// TwinCAT 3 PLC project plc
// ProgramVersion: 3.1.4026.24
// libraries:
//   Tc2_Standard, * (Beckhoff Automation GmbH)
//   Tc2_System, * (Beckhoff Automation GmbH)
//   Tc3_Database, * (Beckhoff Automation GmbH)
// project tree:
//   DUTs/ ST_Signals.TcDUT
//   / PlcTask.TcTTO
//   POUs/ E_FunctionType.TcDUT, FB_FunctionGenerator.TcPOU, MAIN.TcPOU
// real-time tasks:
//   TASK PlcTask: cycle T#10ms, priority 20, ADS port 350

CONFIGURATION plc
    RESOURCE PLC ON TwinCAT3
        TASK PlcTask(INTERVAL := T#10ms, PRIORITY := 20);
        PROGRAM MAIN WITH PlcTask : MAIN;
    END_RESOURCE
END_CONFIGURATION

// ---- DUTs/ST_Signals.TcDUT
TYPE ST_Signals :
STRUCT
    {attribute 'TagName' := 'ID'}
    signal : STRING(255);
    
    {attribute 'FieldName' := 'Value'}
    value : LREAL := -1;
	
END_STRUCT
END_TYPE

// ---- POUs/E_FunctionType.TcDUT
TYPE E_FunctionType :
(
	eSine,
	eSquare,
	ePulse,
	eTriangular,
	eSawtooth,	
	eAM
);
END_TYPE

// ---- POUs/MAIN.TcPOU
PROGRAM MAIN
VAR
	fbSignalSaw				: FB_FunctionGenerator;
	rSignal1				: LREAL;		// Señal dientes de sierra generada por plc
	fbSignalSinus1			: FB_FunctionGenerator;
	rSignal2				: LREAL;		// Señal senoidal generada por plc
	fbDBAutoLog				: FB_PLCDBAutoLogEvt(sNetID:='', tTimeout:=T#5S);
	bAutoLogStart			: BOOL;
	bErrAutoLog				: BOOL;
	aAutoLogStatus			: ARRAY [1..1] OF ST_AutoLogGrpStatus;		// Estado de la conexion Autolog con la DB
	rTrig1					: R_TRIG;
	fTrig2					: F_TRIG;
	bRun					: BOOL;			// Arranca DB Autolog
	bStop					: BOOL;			// Detiene DB Autolog
	timerReset				: TON;
	bErrorInfluxdb			: BOOL;			// Error en la conexion con la DB
	iReconexiones			: INT;			// Contador de reintentos de conexion con la DB
END_VAR

fbSignalSaw(
	bEnable:= TRUE, 
	fFrequency:= 0.2, 
	fAmplitude:= 10, 
	fOffset:= 0, 
	nDutyCycle:= , 
	eFunction:= E_FunctionType.eSawtooth, 
	rSignal:= rSignal1, 
	bError=> );
	
fbSignalSinus1(
	bEnable:= TRUE, 
	fFrequency:= 0.1, 
	fAmplitude:= 5, 
	fOffset:= 0, 
	nDutyCycle:= , 
	eFunction:= E_FunctionType.eSine, 
	rSignal:= rSignal2, 
	bError=> );

rTrig1(CLK:=bAutoLogStart, Q=> );
fTrig2(CLK:=bAutoLogStart, Q=> );

IF _TaskInfo[1].FirstCycle THEN
	bAutoLogStart := TRUE;  // No se inicializa la variable en la declaracion ya que el bloque trigger no detectaría el cambio
END_IF

// Se usa la salida trigger para generar el mensaje en el log, que solo necesita 1 ciclo
// La activacion del autolog con el método Start() tarda unos ciclos
IF rTrig1.Q THEN
	ADSLOGSTR(msgCtrlMask:= ADSLOG_MSGTYPE_WARN OR ADSLOG_MSGTYPE_LOG, msgFmtStr:= 'Autolog Started %s', strArg:='' );
	bRun := TRUE;
END_IF

IF fTrig2.Q THEN
	ADSLOGSTR(msgCtrlMask:= ADSLOG_MSGTYPE_WARN OR ADSLOG_MSGTYPE_LOG, msgFmtStr:= 'Autolog Stopped %s', strArg:='' );
	bStop := TRUE;
END_IF

IF bRun THEN
	IF fbDBAutoLog.Start() THEN
		bRun := FALSE;
	END_IF
END_IF

// EL método Stop también necesita varios ciclos
IF bStop THEN
	IF fbDBAutoLog.Stop() THEN
		bStop := FALSE;
	END_IF
END_IF

// El método de diagnóstico se puede ejecutar cíclicamente
IF bAutoLogStart THEN
	aAutoLogStatus[1].hAutoLogGrpID := 3;
	fbDBAutoLog.Status(tCheckCycle:=T#3S , pError:=ADR(bErrAutoLog) , pAutoLogGrpStatus:=ADR(aAutoLogStatus) , cbAutoLogGrpStatus:=SIZEOF(aAutologStatus) );
	// Si devuelve aAutoLogStatus[1].hrErrorCode= 16#989103E8 la base de datos InfluxDB está detenida
	IF NOT fbDBAutoLog.bBusy_Status THEN
		bErrorInfluxdb := aAutoLogStatus[1].bError;
	END_IF
END_IF

// En caso de error en la conexion con InfluxDB, resetea la funcion autolog cada 3s y comprueba la conexion 
IF bErrorInfluxdb THEN
	bAutoLogStart := FALSE;
	timerReset(IN:=TRUE , PT:=T#3S);
	IF timerReset.Q THEN
		bAutoLogStart := TRUE;
		IF NOT fbDBAutoLog.bBusy_Status THEN
			iReconexiones := iReconexiones+1;
			timerReset(IN:=FALSE);
			bErrorInfluxdb := aAutoLogStatus[1].bError;
		END_IF
	END_IF
ELSE
	timerReset(IN:=FALSE);	
END_IF

END_PROGRAM

// ---- POUs/FB_FunctionGenerator.TcPOU
// Generates a signal build up by the specified function type. v1.2
FUNCTION_BLOCK FB_FunctionGenerator
VAR_INPUT
	bEnable		: BOOL := TRUE;
	fFrequency	: LREAL := 1000;	// in [Hz]
	fAmplitude	: LREAL := 1;
	fOffset		: LREAL;
	nDutyCycle	: UINT := 50;		// % (for pulse function)
	eFunction	: E_FunctionType := E_FunctionType.eSine;	//Default sine wave
END_VAR
VAR_IN_OUT
	rSignal		: LREAL;			//output signal
END_VAR
VAR_OUTPUT
	bError		: BOOL;
END_VAR

VAR
	bInit						: BOOL := TRUE;
	fbGetTaskIdx				: GETCURTASKINDEX;
	
	fLastFrequency				: LREAL;		// in [Hz]
	fLastAmplitude				: LREAL;
	fLastOffset					: LREAL;
	nLastDutyCycle				: UINT;
	eLastFunction				: E_FunctionType;
	
//	nSamples					: UDINT;
	fCycleTime					: LREAL;		// in [s]
	fDelta						: LREAL;		// amplitude delta per sample
	fPhase						: LREAL;		// in [°]
	nSign						: INT := 1;		// 1 or -1
	fLastSignalValue			: LREAL;		// amplitude
	fPeriod						: LREAL;		// in [s]
	fAngularIncrement			: LREAL;		// in [°]
	fAngularIncrementPerCycle	: LREAL;		// in [°]
	fAngularIncrementPerSample	: LREAL;		// in [°]
	(* for modulated signal *)
	fCarrierFrequency			: LREAL := 500;	// in [Hz] (sine)
	fCarrierAmplitude			: LREAL := 1;
	fCarrierPeriod				: LREAL;		// in [s]
	fCarrierAngularIncrement			: LREAL;		// in [°]
	fCarrierAngularIncrementPerCycle	: LREAL;		// in [°]
//	fCarrierAngularIncrementPerSample	: LREAL;		// in [°]
END_VAR

IF bEnable THEN
	IF fLastFrequency <> fFrequency THEN
		bInit := TRUE; // For automatic initializing
		fLastFrequency := fFrequency;
	END_IF
	IF fLastAmplitude <> fAmplitude THEN
		bInit := TRUE; // For automatic initializing
		fLastAmplitude := fAmplitude;
	END_IF
	IF fLastOffset <> fOffset THEN
		bInit := TRUE; // For automatic initializing
		fLastOffset := fOffset;
	END_IF
	IF nLastDutyCycle <> nDutyCycle THEN
		bInit := TRUE; // For automatic initializing
		nLastDutyCycle := nDutyCycle;
	END_IF
	IF eLastFunction <> eFunction THEN
		bInit := TRUE; // For automatic initializing
		eLastFunction := eFunction;
	END_IF
	IF bInit THEN
		// Get taks info	
		fbGetTaskIdx();
		fCycleTime := TwinCAT_SystemInfoVarList._TaskInfo[fbGetTaskIdx.index].CycleTime (*100ns*) / (10.0 * 1000.0 * 1000.0);	
		fLastSignalValue := 0;
		nSign := 1;
		fAngularIncrement := 0;
		// Flush out old data
		MEMSET(ADR(rSignal), 0, SIZEOF(rSignal));
		IF fFrequency <> 0 AND fCycleTime > 0 THEN		
			// Calculate period, increments per plc cycle, increment per oversample

			IF eFunction = E_FunctionType.eSine THEN
				fPeriod := 1/fFrequency;
				fAngularIncrementPerCycle := 360*(fCycleTime/fPeriod);
				// no phase adjustment
				bInit := FALSE;	
			ELSIF eFunction = E_FunctionType.eSquare	THEN
				fPeriod := 1/fFrequency;
				fAngularIncrementPerCycle  := 360*(fCycleTime/fPeriod);
				fPhase := 0.5*360;
				bInit := FALSE;
			ELSIF eFunction = E_FunctionType.ePulse THEN
				fPeriod := 1/fFrequency;
				fAngularIncrementPerCycle  := 360*(fCycleTime/fPeriod);
				IF nDutyCycle > 100 THEN
					nDutyCycle := 100;
				END_IF
				fPhase := (UDINT_TO_LREAL(nDutyCycle)/100)*360;
				bInit := FALSE;					
			ELSIF eFunction = E_FunctionType.eTriangular THEN
				fPeriod := 1/fFrequency;				
				fAngularIncrementPerCycle  := 360*(fCycleTime/fPeriod);
				fAngularIncrementPerSample := fAngularIncrementPerCycle;
				fPhase := 0.5*360; 
				fDelta := 4*(fAmplitude/(360/fAngularIncrementPerSample));				
				bInit := FALSE;
			ELSIF eFunction = E_FunctionType.eSawtooth THEN
				fPeriod := 1/fFrequency;			
				fAngularIncrementPerCycle  := 360*(fCycleTime/fPeriod);		
				fAngularIncrementPerSample := fAngularIncrementPerCycle;
				fDelta := fAmplitude/(360/fAngularIncrementPerSample);
				bInit := FALSE;
			ELSIF eFunction = E_FunctionType.eAM THEN
				fPeriod := 1/fFrequency;
				fAngularIncrementPerCycle := 360*(fCycleTime/fPeriod);
				// no phase adjustment
				fCarrierPeriod := 1/fCarrierFrequency;
				fCarrierAngularIncrementPerCycle := 360*(fCycleTime/fCarrierPeriod);
				// no phase adjustment	
				bInit := FALSE;			
			ELSE
				bError := TRUE;	
			END_IF
		ELSE
			bError := TRUE;
		END_IF
	END_IF
	
	// Enable function generator
	IF NOT bError THEN		
		CASE eFunction OF		
			// sine: typical for vibrations originating from rotating machine
			E_FunctionType.eSine: Sine();
			
			// square: mixed sine signals good for analyzing spectrum				
			E_FunctionType.eSquare: Square();
			
			// pulse: mixed sine signals good for analyzing spectrum				
			E_FunctionType.ePulse: Pulse();
	
			// sawtooth: ramp-type vibrations, continuously increasing			
			E_FunctionType.eSawtooth: Sawtooth();
		
			// triangular: mixed sine signals good for analyzing spectrum
			E_FunctionType.eTriangular: Triangular();
		
			// amplitude modulation: typical for vibrations originating from gear-tooth failure or bearing faults
			// Carrier signal with own frequency and amplitude		
			E_FunctionType.eAM: AM();			
		END_CASE
	END_IF
ELSE
	// Flush out old data
	MEMSET(ADR(rSignal), 0, SIZEOF(rSignal));
END_IF

METHOD PRIVATE AM
VAR_INPUT
END_VAR
// base signal * carrier signal
rSignal:= ( fAmplitude*SIN(2*PI*(fAngularIncrement)/360) + fOffset )
						* ( fCarrierAmplitude*SIN(2*PI*(fCarrierAngularIncrement)/360) );

// Increment angular positions
fAngularIncrement := fAngularIncrement + fAngularIncrementPerCycle;
fCarrierAngularIncrement := fCarrierAngularIncrement + fCarrierAngularIncrementPerCycle;
END_METHOD

METHOD PRIVATE Pulse
VAR_INPUT
END_VAR
// For pulse wave (unequal phases)
IF (fAngularIncrement >= 360) THEN
	fAngularIncrement := fAngularIncrement - DINT_TO_LREAL(LREAL_TO_DINT(fAngularIncrement/360))*360;
	// or with Tc2_Math library: fAngularIncrement := LMOD(fAngularIncrement,360);
END_IF
IF (fAngularIncrement < fPhase) THEN
	nSign := 1;		
ELSIF (fAngularIncrement >= fPhase) THEN
	nSign := 0;
END_IF

rSignal:= nSign*fAmplitude;

rSignal:= rSignal+ fOffset;
END_METHOD

METHOD PRIVATE Sawtooth
VAR_INPUT
END_VAR

// For sawtooth wave (equal phase = period/2)
IF (fAngularIncrement >= 360) THEN
	fAngularIncrement := fAngularIncrement - DINT_TO_LREAL(LREAL_TO_DINT(fAngularIncrement/360))*360;
	// or with Tc2_Math library: fAngularIncrement := LMOD(fAngularIncrement,360);
	fLastSignalValue := fLastSignalValue -fAmplitude;
END_IF
fAngularIncrement := fAngularIncrement + fAngularIncrementPerSample;

rSignal:= fLastSignalValue + fDelta;

// Store last sample
fLastSignalValue := rSignal;

rSignal:= rSignal+ fOffset;
END_METHOD

METHOD PRIVATE Sine
VAR_INPUT
END_VAR

rSignal := fAmplitude*SIN(2*PI*(fAngularIncrement/360));

rSignal := rSignal + fOffset;


// Increment angular position
fAngularIncrement := fAngularIncrement + fAngularIncrementPerCycle;
END_METHOD

METHOD PRIVATE Square
VAR_INPUT
END_VAR

// For square wave (equal phase = period/2)
IF (fAngularIncrement >= 360) THEN
	fAngularIncrement := fAngularIncrement - DINT_TO_LREAL(LREAL_TO_DINT(fAngularIncrement/360))*360;
	// or with Tc2_Math library: fAngularIncrement := LMOD(fAngularIncrement,360);
END_IF
IF (fAngularIncrement < fPhase) THEN
	nSign := 1;
ELSIF (fAngularIncrement >= fPhase) THEN
	nSign := -1;
END_IF

rSignal := nSign*fAmplitude;

rSignal := rSignal + fOffset;
END_METHOD

METHOD PRIVATE Triangular
VAR_INPUT
END_VAR

IF (fAngularIncrement >= 360) THEN
	fAngularIncrement := fAngularIncrement - DINT_TO_LREAL(LREAL_TO_DINT(fAngularIncrement/360))*360;
	// or with Tc2_Math library: fAngularIncrement := LMOD(fAngularIncrement,360);
END_IF
// Negative delta -> Positive delta
IF fAngularIncrement < fPhase/2 THEN	
	nSign := 1;		
ELSIF fAngularIncrement >= fPhase/2 AND fAngularIncrement < 3*fPhase/2 THEN
	nSign := -1;
ELSIF fAngularIncrement >= 3*fPhase/2 THEN
	nSign := 1;	
END_IF
fAngularIncrement := fAngularIncrement + fAngularIncrementPerSample;

rSignal:= fLastSignalValue + nSign*fDelta;
IF rSignal > fAmplitude THEN
	rSignal := rSignal - 2*(rSignal-fAmplitude);
ELSIF rSignal < (-1)*fAmplitude THEN
	rSignal := rSignal - 2*(rSignal+fAmplitude);
END_IF

// Store last sample
fLastSignalValue := rSignal;		

rSignal:= rSignal+ fOffset;
END_METHOD

END_FUNCTION_BLOCK
